Fanuc KAREL source: kt00088.KL

-- PROVISIONAL review KL for V940-1; original PC SHA256 b1fa4f58a401b6a101777f806b09e9d8b727d65e014f72f7aeaab6138734c2ec
-- Incomplete behavior may be omitted. Consult companion uncertainty JSON. Do not deploy.
PROGRAM KT00088
%NOLOCKGROUP
VAR
  OUT : REAL
-- UNRESOLVED_DECL Y1 type=002018
-- UNRESOLVED_DECL H2 type=002017
BEGIN
  -- V9_ZERO_TABLE_METADATA_HINT layout=0001; no indexed target words; source/name/runtime held
  -- UNRESOLVED_PC offsets 5-19; opcodes 2E,22,9D,33,B2
  -- UNRESOLVED_PC offsets 24-38; opcodes 2E,22,9D,33,B4
  -- UNRESOLVED_PC offsets 43-69; opcodes 22,9D,33,B1,22,9D,33,B3,54,64,23
  -- UNRESOLVED_PC offsets 74-78; opcodes 7F
END KT00088
